(* IEC 61131-3 sources: plc-st-coding-agent/progress/evidence/f14_v14_remaining_20261113/jobs/custom_deepseek-v4pro, 30 files *)

(* ---- self-easy-01.candidate_01.st ---- *)
(*
ENGINEERING_CONTRACT
- activation: avgOut updates only when enable=TRUE AND avgEnable=TRUE AND count>0 after clipping count into 1..8.
- hold/retention: enable=FALSE, avgEnable=FALSE, or count<=0 leaves local_avg and avgOut unchanged this scan (S1/S2/S5).
- reset: none specified; avgOut persists until next valid compute; initial local_avg defaults to 0.0.
- boundary: count<=0 causes no division; count>8 uses first 8 samples only (PUB003/PUB004, no overflow).
- precision: sum accumulated in LINT, then converted to REAL and divided by REAL sample count (PUB005/PUB006).
- interface types preserved exactly; no edge-only triggers or interlocks added.
*)

(* CONTRACT_RULES [] *)

FUNCTION_BLOCK FB
VAR_INPUT
    enable: BOOL;
    values: ARRAY[1..8] OF INT;
    count: INT;
    avgEnable: BOOL;
END_VAR
VAR_OUTPUT
    avgOut: REAL;
END_VAR
VAR
    tmp_len: INT;
    tmp_sum: LINT;
    tmp_i: INT;
    local_avg: REAL := 0.0;
END_VAR

IF enable AND avgEnable THEN
    tmp_len := count;
    IF tmp_len < 0 THEN
        tmp_len := 0;
    END_IF;
    IF tmp_len > 8 THEN
        tmp_len := 8;
    END_IF;
    IF tmp_len > 0 THEN
        tmp_sum := 0;
        FOR tmp_i := 1 TO tmp_len BY 1 DO
            tmp_sum := tmp_sum + INT_TO_LINT(values[tmp_i]);
        END_FOR;
        local_avg := LINT_TO_REAL(tmp_sum) / INT_TO_REAL(tmp_len);
    END_IF;
END_IF;

avgOut := local_avg;

END_FUNCTION_BLOCK

(* ---- self-easy-01.raw_candidate_01.st ---- *)
(*
ENGINEERING_CONTRACT
- activation: avgOut updates only when enable=TRUE AND avgEnable=TRUE AND count>0 after clipping count into 1..8.
- hold/retention: enable=FALSE, avgEnable=FALSE, or count<=0 leaves local_avg and avgOut unchanged this scan (S1/S2/S5).
- reset: none specified; avgOut persists until next valid compute; initial local_avg defaults to 0.0.
- boundary: count<=0 causes no division; count>8 uses first 8 samples only (PUB003/PUB004, no overflow).
- precision: sum accumulated in LINT, then converted to REAL and divided by REAL sample count (PUB005/PUB006).
- interface types preserved exactly; no edge-only triggers or interlocks added.
*)

(* CONTRACT_RULES [] *)

FUNCTION_BLOCK FB
VAR_INPUT
    enable: BOOL;
    values: ARRAY[1..8] OF INT;
    count: INT;
    avgEnable: BOOL;
END_VAR
VAR_OUTPUT
    avgOut: REAL;
END_VAR
VAR
    tmp_len: INT;
    tmp_sum: LINT;
    tmp_i: INT;
    local_avg: REAL := 0.0;
END_VAR

IF enable AND avgEnable THEN
    tmp_len := count;
    IF tmp_len < 0 THEN
        tmp_len := 0;
    END_IF;
    IF tmp_len > 8 THEN
        tmp_len := 8;
    END_IF;
    IF tmp_len > 0 THEN
        tmp_sum := 0;
        FOR tmp_i := 1 TO tmp_len BY 1 DO
            tmp_sum := tmp_sum + INT_TO_LINT(values[tmp_i]);
        END_FOR;
        local_avg := LINT_TO_REAL(tmp_sum) / INT_TO_REAL(tmp_len);
    END_IF;
END_IF;

avgOut := local_avg;

END_FUNCTION_BLOCK

(* ---- self-easy-02.candidate_01.st ---- *)
FUNCTION_BLOCK FB
VAR_INPUT
    tankLevel : REAL;
    outletFlow : REAL;
    inletPermit : BOOL;
    resetBtn : BOOL;
END_VAR
VAR_OUTPUT
    pumpRun : BOOL;
    alarmHigh : BOOL;
    alarmLow : BOOL;
    outletValveOpen : BOOL;
END_VAR
VAR
    highLatched : BOOL := FALSE;
    lowLatched : BOOL := FALSE;
    prevResetBtn : BOOL := FALSE;
    tmp_resetRising : BOOL;
END_VAR

(* ENGINEERING_CONTRACT
   alarmHigh/alarmLow: set immediately at respective threshold, then latch.
   Activation: high >= 85.0, low <= 15.0 (REAL percent).
   Retention: remain latched when level returns to normal until reset.
   Reset: resetBtn rising edge clears each latch only if its danger is absent.
   Same-scan priority: danger condition overrides reset for the affected alarm.
   pumpRun: active only when inletPermit AND no alarm latched.
   outletValveOpen: inverse of low alarm; outletFlow is unused observation input.
*)

(* CONTRACT_RULES [] *)

tmp_resetRising := resetBtn AND NOT prevResetBtn;

IF tankLevel >= 85.0 THEN
    highLatched := TRUE;
ELSIF tmp_resetRising THEN
    highLatched := FALSE;
END_IF;

IF tankLevel <= 15.0 THEN
    lowLatched := TRUE;
ELSIF tmp_resetRising THEN
    lowLatched := FALSE;
END_IF;

alarmHigh := highLatched;
alarmLow := lowLatched;
pumpRun := inletPermit AND NOT highLatched AND NOT lowLatched;
outletValveOpen := NOT lowLatched;

prevResetBtn := resetBtn;

END_FUNCTION_BLOCK

(* ---- self-easy-02.raw_candidate_01.st ---- *)
FUNCTION_BLOCK FB
VAR_INPUT
    tankLevel : REAL;
    outletFlow : REAL;
    inletPermit : BOOL;
    resetBtn : BOOL;
END_VAR
VAR_OUTPUT
    pumpRun : BOOL;
    alarmHigh : BOOL;
    alarmLow : BOOL;
    outletValveOpen : BOOL;
END_VAR
VAR
    highLatched : BOOL := FALSE;
    lowLatched : BOOL := FALSE;
    prevResetBtn : BOOL := FALSE;
    tmp_resetRising : BOOL;
END_VAR

(* ENGINEERING_CONTRACT
   alarmHigh/alarmLow: set immediately at respective threshold, then latch.
   Activation: high >= 85.0, low <= 15.0 (REAL percent).
   Retention: remain latched when level returns to normal until reset.
   Reset: resetBtn rising edge clears each latch only if its danger is absent.
   Same-scan priority: danger condition overrides reset for the affected alarm.
   pumpRun: active only when inletPermit AND no alarm latched.
   outletValveOpen: inverse of low alarm; outletFlow is unused observation input.
*)

(* CONTRACT_RULES [] *)

tmp_resetRising := resetBtn AND NOT prevResetBtn;

IF tankLevel >= 85.0 THEN
    highLatched := TRUE;
ELSIF tmp_resetRising THEN
    highLatched := FALSE;
END_IF;

IF tankLevel <= 15.0 THEN
    lowLatched := TRUE;
ELSIF tmp_resetRising THEN
    lowLatched := FALSE;
END_IF;

alarmHigh := highLatched;
alarmLow := lowLatched;
pumpRun := inletPermit AND NOT highLatched AND NOT lowLatched;
outletValveOpen := NOT lowLatched;

prevResetBtn := resetBtn;

END_FUNCTION_BLOCK

(* ---- self-hard-01.candidate_01.st ---- *)
(*
ENGINEERING_CONTRACT
alarmActive: next = flowLow OR (prevActive AND !risingAck AND !(prevFlowLow AND prevAcked)).
  Retain on unacked condition loss; clear only when active-acked and flowLow drops, or ack rising while flowLow false.
alarmAcked: next = nextActive AND (!flowLow OR risingAck OR (prevFlowLow AND prevActive AND prevAcked)).
  True for active/acked or pending-clear; false when inactive or new flowLow after pending-clear.
highHigh = NOT sensorOK (combinational; no latch; auto clears same scan as sensorOK).
Memory: prevFlowLow/prevActive/prevAcked/prevAckBtn retained in VAR; update after output assignment.
Same-scan: risingAck computed before outputs; formulas use previous-cycle stored state; high priority independent.
Units: BOOL; no timers. See PUB001-PUB038.
*)
(* CONTRACT_RULES [] *)
FUNCTION_BLOCK FB
VAR_INPUT
    flowLow: BOOL;
    ackBtn: BOOL;
    sensorOK: BOOL;
END_VAR
VAR_OUTPUT
    alarmActive: BOOL;
    alarmAcked: BOOL;
    highHigh: BOOL;
END_VAR
VAR
    prevFlowLow: BOOL;
    prevAlarmActive: BOOL;
    prevAlarmAcked: BOOL;
    prevAckBtn: BOOL;
    risingAck: BOOL;
    nextActive: BOOL;
    nextAcked: BOOL;
    prevFlowLowAndAcked: BOOL;
    prevFlowLowActiveAcked: BOOL;
END_VAR

risingAck := ackBtn AND NOT prevAckBtn;

prevFlowLowAndAcked := prevFlowLow AND prevAlarmAcked;
prevFlowLowActiveAcked := prevFlowLow AND prevAlarmActive AND prevAlarmAcked;

nextActive := flowLow OR (prevAlarmActive AND NOT risingAck AND (NOT prevFlowLowAndAcked));
nextAcked := nextActive AND (NOT flowLow OR risingAck OR prevFlowLowActiveAcked);

alarmActive := nextActive;
alarmAcked := nextAcked;
highHigh := NOT sensorOK;

prevFlowLow := flowLow;
prevAlarmActive := nextActive;
prevAlarmAcked := nextAcked;
prevAckBtn := ackBtn;

END_FUNCTION_BLOCK

(* ---- self-hard-01.raw_candidate_01.st ---- *)
(*
ENGINEERING_CONTRACT
alarmActive: next = flowLow OR (prevActive AND !risingAck AND !(prevFlowLow AND prevAcked)).
  Retain on unacked condition loss; clear only when active-acked and flowLow drops, or ack rising while flowLow false.
alarmAcked: next = nextActive AND (!flowLow OR risingAck OR (prevFlowLow AND prevActive AND prevAcked)).
  True for active/acked or pending-clear; false when inactive or new flowLow after pending-clear.
highHigh = NOT sensorOK (combinational; no latch; auto clears same scan as sensorOK).
Memory: prevFlowLow/prevActive/prevAcked/prevAckBtn retained in VAR; update after output assignment.
Same-scan: risingAck computed before outputs; formulas use previous-cycle stored state; high priority independent.
Units: BOOL; no timers. See PUB001-PUB038.
*)
(* CONTRACT_RULES [] *)
FUNCTION_BLOCK FB
VAR_INPUT
    flowLow: BOOL;
    ackBtn: BOOL;
    sensorOK: BOOL;
END_VAR
VAR_OUTPUT
    alarmActive: BOOL;
    alarmAcked: BOOL;
    highHigh: BOOL;
END_VAR
VAR
    prevFlowLow: BOOL;
    prevAlarmActive: BOOL;
    prevAlarmAcked: BOOL;
    prevAckBtn: BOOL;
    risingAck: BOOL;
    nextActive: BOOL;
    nextAcked: BOOL;
    prevFlowLowAndAcked: BOOL;
    prevFlowLowActiveAcked: BOOL;
END_VAR

risingAck := ackBtn AND NOT prevAckBtn;

prevFlowLowAndAcked := prevFlowLow AND prevAlarmAcked;
prevFlowLowActiveAcked := prevFlowLow AND prevAlarmActive AND prevAlarmAcked;

nextActive := flowLow OR (prevAlarmActive AND NOT risingAck AND (NOT prevFlowLowAndAcked));
nextAcked := nextActive AND (NOT flowLow OR risingAck OR prevFlowLowActiveAcked);

alarmActive := nextActive;
alarmAcked := nextAcked;
highHigh := NOT sensorOK;

prevFlowLow := flowLow;
prevAlarmActive := nextActive;
prevAlarmAcked := nextAcked;
prevAckBtn := ackBtn;

END_FUNCTION_BLOCK

(* ---- self-hard-02.candidate_01.st ---- *)
FUNCTION_BLOCK FB
VAR_INPUT
    startBtn : BOOL;
    abortBtn : BOOL;
    setpoint : REAL;
    pv : REAL;
    maxDuration : INT;
END_VAR
VAR_OUTPUT
    elapsed : INT;
    phase : INT;
    timeout : BOOL;
END_VAR
VAR
    prevStartBtn : BOOL;
    tmpStartRising : BOOL;
    tmpPrevPhase : INT;
    tmpPrevElapsed : INT;
    tmpPrevTimeout : BOOL;
    tmpIsRunPrev : BOOL;
    tmpNewElapsed : INT;
END_VAR

(* ENGINEERING_CONTRACT
   phase: 0 idle, 1 heating, 2 soaking, 3 done, 9 aborted.
   Activation: phase=1 on start rising without abort; phase=2 when previous run phase is 1 and pv>=setpoint before timeout; phase=3 when elapsed>=maxDuration; phase=9 on abort.
   Retention: phase 3/9 hold until new start or abort; start resets to 1 and clears elapsed/timeout; abort from 3/9 preserves elapsed/timeout.
   elapsed: counts scans when previous phase is 1 or 2 and no abort/start rising. Reset to 0 on start; frozen in 3/9; frozen on abort.
   timeout: set TRUE when new elapsed>=maxDuration (scan count); cleared on start; frozen on abort; otherwise equals timeout condition.
   Priority: abort > start rising > running count; same-scan start edge consumed even under abort.
   Units: elapsed/maxDuration in scan counts, INT; no timer used.
*)

(* CONTRACT_RULES [] *)

tmpStartRising := startBtn AND NOT prevStartBtn;
tmpPrevPhase := phase;
tmpPrevElapsed := elapsed;
tmpPrevTimeout := timeout;
tmpIsRunPrev := (tmpPrevPhase = 1) OR (tmpPrevPhase = 2);

IF abortBtn THEN
    phase := 9;
    elapsed := tmpPrevElapsed;
    timeout := tmpPrevTimeout;
ELSIF tmpStartRising THEN
    phase := 1;
    elapsed := 0;
    timeout := FALSE;
ELSE
    IF tmpIsRunPrev THEN
        tmpNewElapsed := tmpPrevElapsed + 1;
        elapsed := tmpNewElapsed;
        IF tmpNewElapsed >= maxDuration THEN
            timeout := TRUE;
            phase := 3;
        ELSE
            timeout := FALSE;
            IF tmpPrevPhase = 2 THEN
                phase := 2;
            ELSE
                IF pv >= setpoint THEN
                    phase := 2;
                ELSE
                    phase := 1;
                END_IF;
            END_IF;
        END_IF;
    ELSE
        phase := tmpPrevPhase;
        elapsed := tmpPrevElapsed;
        timeout := tmpPrevTimeout;
    END_IF;
END_IF;

prevStartBtn := startBtn;
END_FUNCTION_BLOCK

(* ---- self-hard-02.raw_candidate_01.st ---- *)
FUNCTION_BLOCK FB
VAR_INPUT
    startBtn : BOOL;
    abortBtn : BOOL;
    setpoint : REAL;
    pv : REAL;
    maxDuration : INT;
END_VAR
VAR_OUTPUT
    elapsed : INT;
    phase : INT;
    timeout : BOOL;
END_VAR
VAR
    prevStartBtn : BOOL;
    tmpStartRising : BOOL;
    tmpPrevPhase : INT;
    tmpPrevElapsed : INT;
    tmpPrevTimeout : BOOL;
    tmpIsRunPrev : BOOL;
    tmpNewElapsed : INT;
END_VAR

(* ENGINEERING_CONTRACT
   phase: 0 idle, 1 heating, 2 soaking, 3 done, 9 aborted.
   Activation: phase=1 on start rising without abort; phase=2 when previous run phase is 1 and pv>=setpoint before timeout; phase=3 when elapsed>=maxDuration; phase=9 on abort.
   Retention: phase 3/9 hold until new start or abort; start resets to 1 and clears elapsed/timeout; abort from 3/9 preserves elapsed/timeout.
   elapsed: counts scans when previous phase is 1 or 2 and no abort/start rising. Reset to 0 on start; frozen in 3/9; frozen on abort.
   timeout: set TRUE when new elapsed>=maxDuration (scan count); cleared on start; frozen on abort; otherwise equals timeout condition.
   Priority: abort > start rising > running count; same-scan start edge consumed even under abort.
   Units: elapsed/maxDuration in scan counts, INT; no timer used.
*)

(* CONTRACT_RULES [] *)

tmpStartRising := startBtn AND NOT prevStartBtn;
tmpPrevPhase := phase;
tmpPrevElapsed := elapsed;
tmpPrevTimeout := timeout;
tmpIsRunPrev := (tmpPrevPhase = 1) OR (tmpPrevPhase = 2);

IF abortBtn THEN
    phase := 9;
    elapsed := tmpPrevElapsed;
    timeout := tmpPrevTimeout;
ELSIF tmpStartRising THEN
    phase := 1;
    elapsed := 0;
    timeout := FALSE;
ELSE
    IF tmpIsRunPrev THEN
        tmpNewElapsed := tmpPrevElapsed + 1;
        elapsed := tmpNewElapsed;
        IF tmpNewElapsed >= maxDuration THEN
            timeout := TRUE;
            phase := 3;
        ELSE
            timeout := FALSE;
            IF tmpPrevPhase = 2 THEN
                phase := 2;
            ELSE
                IF pv >= setpoint THEN
                    phase := 2;
                ELSE
                    phase := 1;
                END_IF;
            END_IF;
        END_IF;
    ELSE
        phase := tmpPrevPhase;
        elapsed := tmpPrevElapsed;
        timeout := tmpPrevTimeout;
    END_IF;
END_IF;

prevStartBtn := startBtn;
END_FUNCTION_BLOCK

(* ---- self-hard-03.candidate_01.st ---- *)
(* ENGINEERING_CONTRACT
   count: updated by successful pop then successful push; retained otherwise; initial 0; bounds 0..8; S1,S6.
   full: combinational = (count=8); no latch; S1.
   empty: combinational = (count=0); no latch; S1.
   head: count=0 -> 0; else fifo[1]; combinational after actions; S5.
   fifo valid prefix: compact; shift on successful pop; append on successful push; S4,S7,S8.
   Edge history: local_push_prev/local_pop_prev retained; initial FALSE; updated each scan.
   Priority: pop rising executes before push rising; capacity checked after pop; PUB requirement order.
*)
(* CONTRACT_RULES [] *)
FUNCTION_BLOCK FB
VAR_INPUT
    pushEn : BOOL;
    pushItem : INT;
    popEn : BOOL;
END_VAR
VAR_OUTPUT
    count : INT;
    full : BOOL;
    empty : BOOL;
    head : INT;
END_VAR
VAR_IN_OUT
    fifo : ARRAY[1..8] OF INT;
END_VAR
VAR
    local_push_prev : BOOL := FALSE;
    local_pop_prev : BOOL := FALSE;
    local_count : INT := 0;
    local_rising_push : BOOL;
    local_rising_pop : BOOL;
    i : INT;
END_VAR

(* 计算上升沿，历史在扫描结束时更新 *)
local_rising_push := pushEn AND NOT local_push_prev;
local_rising_pop := popEn AND NOT local_pop_prev;

(* 先执行出队 *)
IF local_rising_pop AND (local_count > 0) THEN
    IF local_count > 1 THEN
        FOR i := 1 TO local_count - 1 DO
            fifo[i] := fifo[i + 1];
        END_FOR;
    END_IF;
    local_count := local_count - 1;
END_IF;

(* 后执行入队 *)
IF local_rising_push AND (local_count < 8) THEN
    local_count := local_count + 1;
    fifo[local_count] := pushItem;
END_IF;

(* 输出 *)
count := local_count;
full := (local_count = 8);
empty := (local_count = 0);
IF local_count = 0 THEN
    head := 0;
ELSE
    head := fifo[1];
END_IF;

(* 更新输入历史 *)
local_push_prev := pushEn;
local_pop_prev := popEn;

END_FUNCTION_BLOCK

(* ---- self-hard-03.raw_candidate_01.st ---- *)
(* ENGINEERING_CONTRACT
   count: updated by successful pop then successful push; retained otherwise; initial 0; bounds 0..8; S1,S6.
   full: combinational = (count=8); no latch; S1.
   empty: combinational = (count=0); no latch; S1.
   head: count=0 -> 0; else fifo[1]; combinational after actions; S5.
   fifo valid prefix: compact; shift on successful pop; append on successful push; S4,S7,S8.
   Edge history: local_push_prev/local_pop_prev retained; initial FALSE; updated each scan.
   Priority: pop rising executes before push rising; capacity checked after pop; PUB requirement order.
*)
(* CONTRACT_RULES [] *)
FUNCTION_BLOCK FB
VAR_INPUT
    pushEn : BOOL;
    pushItem : INT;
    popEn : BOOL;
END_VAR
VAR_OUTPUT
    count : INT;
    full : BOOL;
    empty : BOOL;
    head : INT;
END_VAR
VAR_IN_OUT
    fifo : ARRAY[1..8] OF INT;
END_VAR
VAR
    local_push_prev : BOOL := FALSE;
    local_pop_prev : BOOL := FALSE;
    local_count : INT := 0;
    local_rising_push : BOOL;
    local_rising_pop : BOOL;
    i : INT;
END_VAR

(* 计算上升沿，历史在扫描结束时更新 *)
local_rising_push := pushEn AND NOT local_push_prev;
local_rising_pop := popEn AND NOT local_pop_prev;

(* 先执行出队 *)
IF local_rising_pop AND (local_count > 0) THEN
    IF local_count > 1 THEN
        FOR i := 1 TO local_count - 1 DO
            fifo[i] := fifo[i + 1];
        END_FOR;
    END_IF;
    local_count := local_count - 1;
END_IF;

(* 后执行入队 *)
IF local_rising_push AND (local_count < 8) THEN
    local_count := local_count + 1;
    fifo[local_count] := pushItem;
END_IF;

(* 输出 *)
count := local_count;
full := (local_count = 8);
empty := (local_count = 0);
IF local_count = 0 THEN
    head := 0;
ELSE
    head := fifo[1];
END_IF;

(* 更新输入历史 *)
local_push_prev := pushEn;
local_pop_prev := popEn;

END_FUNCTION_BLOCK

(* ---- self-hard-04.candidate_01.st ---- *)
(* ENGINEERING_CONTRACT
  runningCount: combinational; activation every scan; clip demand to 0..5; no retention/reset; same-scan priority: computed first; range 0..5 [PUB001,S1].
  leadPump: stored selection; activation: positive demand with prevLead=0 -> global (hours,pump) min (tie smallest pump); positive prevLead valid + rotated TRUE and oldLeadHours-globalMinHours > 50 -> global min; else retain; deactivation/reset: demand<=0 -> 0; units 1..5,0=none [PUB004,S2,S3,S6,S7].
  lagPump: stored selection; activation/update: demand>=2 and (lead changed OR clipped demand rose) -> min among pumps excluding current lead (tie smallest pump); retention: otherwise while demand>=2; deactivation/reset: demand<=1 -> 0; units 1..5,0=none [PUB005,S8,S9].
  Arrays accessed with indices 1..5 only; previous outputs kept in static VAR [PUB006].
*)
(* CONTRACT_RULES [] *)
FUNCTION_BLOCK FB
VAR_INPUT
    demand : INT;
    runHours : ARRAY[1..5] OF LINT;
    rotated : BOOL;
END_VAR
VAR_OUTPUT
    leadPump : INT;
    lagPump : INT;
    runningCount : INT;
END_VAR
VAR
    local_prevLeadPump : INT := 0;
    local_prevLagPump : INT := 0;
    local_prevRunningCount : INT := 0;
    local_demandClipped : INT;
    local_i : INT;
    local_minPumpAll : INT;
    local_minHoursAll : LINT;
    local_minPumpExcl : INT;
    local_minHoursExcl : LINT;
    local_firstFound : BOOL;
END_VAR

IF demand < 0 THEN
    local_demandClipped := 0;
ELSIF demand > 5 THEN
    local_demandClipped := 5;
ELSE
    local_demandClipped := demand;
END_IF;

runningCount := local_demandClipped;

IF local_demandClipped <= 0 THEN
    leadPump := 0;
    lagPump := 0;
ELSE
    local_minPumpAll := 1;
    local_minHoursAll := runHours[1];
    FOR local_i := 2 TO 5 DO
        IF (runHours[local_i] < local_minHoursAll) OR
           ((runHours[local_i] = local_minHoursAll) AND (local_i < local_minPumpAll)) THEN
            local_minPumpAll := local_i;
            local_minHoursAll := runHours[local_i];
        END_IF;
    END_FOR;

    IF local_prevLeadPump = 0 THEN
        leadPump := local_minPumpAll;
    ELSE
        leadPump := local_prevLeadPump;
        IF rotated THEN
            IF runHours[local_prevLeadPump] - local_minHoursAll > LINT#50 THEN
                leadPump := local_minPumpAll;
            END_IF;
        END_IF;
    END_IF;

    IF local_demandClipped = 1 THEN
        lagPump := 0;
    ELSE
        IF (leadPump <> local_prevLeadPump) OR (local_demandClipped > local_prevRunningCount) THEN
            local_minPumpExcl := 0;
            local_minHoursExcl := 0;
            local_firstFound := FALSE;
            FOR local_i := 1 TO 5 DO
                IF local_i <> leadPump THEN
                    IF NOT local_firstFound THEN
                        local_minPumpExcl := local_i;
                        local_minHoursExcl := runHours[local_i];
                        local_firstFound := TRUE;
                    ELSE
                        IF (runHours[local_i] < local_minHoursExcl) OR
                           ((runHours[local_i] = local_minHoursExcl) AND (local_i < local_minPumpExcl)) THEN
                            local_minPumpExcl := local_i;
                            local_minHoursExcl := runHours[local_i];
                        END_IF;
                    END_IF;
                END_IF;
            END_FOR;
            lagPump := local_minPumpExcl;
        ELSE
            lagPump := local_prevLagPump;
        END_IF;
    END_IF;
END_IF;

local_prevLeadPump := leadPump;
local_prevLagPump := lagPump;
local_prevRunningCount := runningCount;

END_FUNCTION_BLOCK

(* ---- self-hard-04.raw_candidate_01.st ---- *)
(* ENGINEERING_CONTRACT
  runningCount: combinational; activation every scan; clip demand to 0..5; no retention/reset; same-scan priority: computed first; range 0..5 [PUB001,S1].
  leadPump: stored selection; activation: positive demand with prevLead=0 -> global (hours,pump) min (tie smallest pump); positive prevLead valid + rotated TRUE and oldLeadHours-globalMinHours > 50 -> global min; else retain; deactivation/reset: demand<=0 -> 0; units 1..5,0=none [PUB004,S2,S3,S6,S7].
  lagPump: stored selection; activation/update: demand>=2 and (lead changed OR clipped demand rose) -> min among pumps excluding current lead (tie smallest pump); retention: otherwise while demand>=2; deactivation/reset: demand<=1 -> 0; units 1..5,0=none [PUB005,S8,S9].
  Arrays accessed with indices 1..5 only; previous outputs kept in static VAR [PUB006].
*)
(* CONTRACT_RULES [] *)
FUNCTION_BLOCK FB
VAR_INPUT
    demand : INT;
    runHours : ARRAY[1..5] OF LINT;
    rotated : BOOL;
END_VAR
VAR_OUTPUT
    leadPump : INT;
    lagPump : INT;
    runningCount : INT;
END_VAR
VAR
    local_prevLeadPump : INT := 0;
    local_prevLagPump : INT := 0;
    local_prevRunningCount : INT := 0;
    local_demandClipped : INT;
    local_i : INT;
    local_minPumpAll : INT;
    local_minHoursAll : LINT;
    local_minPumpExcl : INT;
    local_minHoursExcl : LINT;
    local_firstFound : BOOL;
END_VAR

IF demand < 0 THEN
    local_demandClipped := 0;
ELSIF demand > 5 THEN
    local_demandClipped := 5;
ELSE
    local_demandClipped := demand;
END_IF;

runningCount := local_demandClipped;

IF local_demandClipped <= 0 THEN
    leadPump := 0;
    lagPump := 0;
ELSE
    local_minPumpAll := 1;
    local_minHoursAll := runHours[1];
    FOR local_i := 2 TO 5 DO
        IF (runHours[local_i] < local_minHoursAll) OR
           ((runHours[local_i] = local_minHoursAll) AND (local_i < local_minPumpAll)) THEN
            local_minPumpAll := local_i;
            local_minHoursAll := runHours[local_i];
        END_IF;
    END_FOR;

    IF local_prevLeadPump = 0 THEN
        leadPump := local_minPumpAll;
    ELSE
        leadPump := local_prevLeadPump;
        IF rotated THEN
            IF runHours[local_prevLeadPump] - local_minHoursAll > LINT#50 THEN
                leadPump := local_minPumpAll;
            END_IF;
        END_IF;
    END_IF;

    IF local_demandClipped = 1 THEN
        lagPump := 0;
    ELSE
        IF (leadPump <> local_prevLeadPump) OR (local_demandClipped > local_prevRunningCount) THEN
            local_minPumpExcl := 0;
            local_minHoursExcl := 0;
            local_firstFound := FALSE;
            FOR local_i := 1 TO 5 DO
                IF local_i <> leadPump THEN
                    IF NOT local_firstFound THEN
                        local_minPumpExcl := local_i;
                        local_minHoursExcl := runHours[local_i];
                        local_firstFound := TRUE;
                    ELSE
                        IF (runHours[local_i] < local_minHoursExcl) OR
                           ((runHours[local_i] = local_minHoursExcl) AND (local_i < local_minPumpExcl)) THEN
                            local_minPumpExcl := local_i;
                            local_minHoursExcl := runHours[local_i];
                        END_IF;
                    END_IF;
                END_IF;
            END_FOR;
            lagPump := local_minPumpExcl;
        ELSE
            lagPump := local_prevLagPump;
        END_IF;
    END_IF;
END_IF;

local_prevLeadPump := leadPump;
local_prevLagPump := lagPump;
local_prevRunningCount := runningCount;

END_FUNCTION_BLOCK

(* ---- self-hard-05.candidate_01.st ---- *)
(* ENGINEERING_CONTRACT
tripLatched: set same scan when runRequest=TRUE AND flameOK=FALSE; held; clear only on rising resetBtn while runRequest=FALSE AND flameOK=FALSE; fire-set dominates. PUB001 PUB006 PUB030 PUB031 PUB059.
fuelPermit: combinational = runRequest AND flameOK AND NOT tripLatched. PUB005 PUB060.
o2Fault: combinational = NOT o2Valid OR o2PV<0.0 OR o2PV>21.0. PUB012 PUB061.
trimEnable: combinational = fuelPermit AND NOT o2Fault. PUB008 PUB061.
airTrim: if trimEnable then clamp(2.0*(2.0-o2PV), -10.0, 10.0) else 0.0; saturation reaches -10 only when o2PV>7.0. PUB010 PUB011 PUB014 PUB015 PUB052 PUB053.
airCommand: if fuelPermit then clamp(baseAir+airTrim, 0.0, 100.0) else 0.0. PUB011 PUB013 PUB015 PUB045 PUB046 PUB055.
reset edge: detected once per scan via prevResetBtn; no timer. Units: REAL %, BOOL, scan cycle. PUB006 PUB030 PUB031.
*)
(* CONTRACT_RULES [] *)
FUNCTION_BLOCK FB
VAR_INPUT
    runRequest : BOOL;
    flameOK : BOOL;
    o2Valid : BOOL;
    o2PV : REAL;
    baseAir : REAL;
    resetBtn : BOOL;
END_VAR
VAR_OUTPUT
    fuelPermit : BOOL;
    trimEnable : BOOL;
    airTrim : REAL;
    airCommand : REAL;
    tripLatched : BOOL;
    o2Fault : BOOL;
END_VAR
VAR
    prevResetBtn : BOOL := FALSE;
    tmp_resetRise : BOOL;
    tmp_prevTrip : BOOL;
    tmp_rawTrim : REAL;
    tmp_sum : REAL;
END_VAR

    tmp_resetRise := resetBtn AND NOT prevResetBtn;
    tmp_prevTrip := tripLatched;
    tripLatched := (runRequest AND NOT flameOK)
                   OR (tmp_prevTrip AND NOT (tmp_resetRise AND NOT runRequest AND NOT flameOK));
    prevResetBtn := resetBtn;

    fuelPermit := runRequest AND flameOK AND NOT tripLatched;

    o2Fault := (NOT o2Valid) OR (o2PV < 0.0) OR (o2PV > 21.0);
    trimEnable := fuelPermit AND NOT o2Fault;

    IF trimEnable THEN
        tmp_rawTrim := 2.0 * (2.0 - o2PV);
        IF tmp_rawTrim < -10.0 THEN
            airTrim := -10.0;
        ELSIF tmp_rawTrim > 10.0 THEN
            airTrim := 10.0;
        ELSE
            airTrim := tmp_rawTrim;
        END_IF;
    ELSE
        airTrim := 0.0;
    END_IF;

    IF fuelPermit THEN
        tmp_sum := baseAir + airTrim;
        IF tmp_sum < 0.0 THEN
            airCommand := 0.0;
        ELSIF tmp_sum > 100.0 THEN
            airCommand := 100.0;
        ELSE
            airCommand := tmp_sum;
        END_IF;
    ELSE
        airCommand := 0.0;
    END_IF;

END_FUNCTION_BLOCK

(* ---- self-hard-05.raw_candidate_01.st ---- *)
(* ENGINEERING_CONTRACT
tripLatched: set same scan when runRequest=TRUE AND flameOK=FALSE; held; clear only on rising resetBtn while runRequest=FALSE AND flameOK=FALSE; fire-set dominates. PUB001 PUB006 PUB030 PUB031 PUB059.
fuelPermit: combinational = runRequest AND flameOK AND NOT tripLatched. PUB005 PUB060.
o2Fault: combinational = NOT o2Valid OR o2PV<0.0 OR o2PV>21.0. PUB012 PUB061.
trimEnable: combinational = fuelPermit AND NOT o2Fault. PUB008 PUB061.
airTrim: if trimEnable then clamp(2.0*(2.0-o2PV), -10.0, 10.0) else 0.0; saturation reaches -10 only when o2PV>7.0. PUB010 PUB011 PUB014 PUB015 PUB052 PUB053.
airCommand: if fuelPermit then clamp(baseAir+airTrim, 0.0, 100.0) else 0.0. PUB011 PUB013 PUB015 PUB045 PUB046 PUB055.
reset edge: detected once per scan via prevResetBtn; no timer. Units: REAL %, BOOL, scan cycle. PUB006 PUB030 PUB031.
*)
(* CONTRACT_RULES [] *)
FUNCTION_BLOCK FB
VAR_INPUT
    runRequest : BOOL;
    flameOK : BOOL;
    o2Valid : BOOL;
    o2PV : REAL;
    baseAir : REAL;
    resetBtn : BOOL;
END_VAR
VAR_OUTPUT
    fuelPermit : BOOL;
    trimEnable : BOOL;
    airTrim : REAL;
    airCommand : REAL;
    tripLatched : BOOL;
    o2Fault : BOOL;
END_VAR
VAR
    prevResetBtn : BOOL := FALSE;
    tmp_resetRise : BOOL;
    tmp_prevTrip : BOOL;
    tmp_rawTrim : REAL;
    tmp_sum : REAL;
END_VAR

    tmp_resetRise := resetBtn AND NOT prevResetBtn;
    tmp_prevTrip := tripLatched;
    tripLatched := (runRequest AND NOT flameOK)
                   OR (tmp_prevTrip AND NOT (tmp_resetRise AND NOT runRequest AND NOT flameOK));
    prevResetBtn := resetBtn;

    fuelPermit := runRequest AND flameOK AND NOT tripLatched;

    o2Fault := (NOT o2Valid) OR (o2PV < 0.0) OR (o2PV > 21.0);
    trimEnable := fuelPermit AND NOT o2Fault;

    IF trimEnable THEN
        tmp_rawTrim := 2.0 * (2.0 - o2PV);
        IF tmp_rawTrim < -10.0 THEN
            airTrim := -10.0;
        ELSIF tmp_rawTrim > 10.0 THEN
            airTrim := 10.0;
        ELSE
            airTrim := tmp_rawTrim;
        END_IF;
    ELSE
        airTrim := 0.0;
    END_IF;

    IF fuelPermit THEN
        tmp_sum := baseAir + airTrim;
        IF tmp_sum < 0.0 THEN
            airCommand := 0.0;
        ELSIF tmp_sum > 100.0 THEN
            airCommand := 100.0;
        ELSE
            airCommand := tmp_sum;
        END_IF;
    ELSE
        airCommand := 0.0;
    END_IF;

END_FUNCTION_BLOCK

(* ---- self-hard-06.candidate_01.st ---- *)
(* ENGINEERING_CONTRACT
  tripLatched: active same scan on trip condition (run & !pressureValid) OR (run & pressureValid & pressure>=4500.0);
               retains until legal reset edge: resetBtn rising & !run & pressureValid & pressure<=4200.0.
  fuelPermit: combinational = run & !tripLatched, evaluated after latch update.
  currentCauseMask: low nibble recalculated each scan; !run=0, invalid=1, valid overpressure evaluates stuck/excess/unlocated, below 4500=0.
  latchedCauseMask: OR currentCauseMask while tripLatched; clear when !tripLatched; low 4 bits only.
  stuckCounter: counts consecutive full overpressure+valve-condition scans; reset on any interruption.
  diagnosticActive: currentCauseMask<>0.
  Unspecified: scan period undefined; initial resetBtn edge state considered FALSE.
*)
(* CONTRACT_RULES [] *)
FUNCTION_BLOCK FB
VAR_INPUT
    runRequest : BOOL;
    pressure : REAL;
    pressureValid : BOOL;
    fuelFlow : REAL;
    steamFlow : REAL;
    outletCmd : INT;
    outletFeedback : INT;
    resetBtn : BOOL;
END_VAR
VAR_OUTPUT
    tripLatched : BOOL;
    fuelPermit : BOOL;
    currentCauseMask : WORD;
    latchedCauseMask : WORD;
    diagnosticActive : BOOL;
END_VAR
VAR
    lastResetBtn : BOOL := FALSE;
    stuckCounter : INT := 0;
    tmp_resetRising : BOOL;
    tmp_overpressure : BOOL;
    tmp_invalid : BOOL;
    tmp_tripCondition : BOOL;
    tmp_legalReset : BOOL;
    tmp_stuckCond : BOOL;
    tmp_stuckBit : BOOL;
    tmp_excessBit : BOOL;
END_VAR

tmp_resetRising := resetBtn AND NOT lastResetBtn;
lastResetBtn := resetBtn;

tmp_overpressure := runRequest AND pressureValid AND pressure >= 4500.0;
tmp_invalid := runRequest AND NOT pressureValid;
tmp_tripCondition := tmp_overpressure OR tmp_invalid;
tmp_legalReset := tmp_resetRising AND NOT runRequest AND pressureValid AND pressure <= 4200.0;

IF NOT runRequest THEN
    currentCauseMask := WORD#0;
    stuckCounter := 0;
ELSIF NOT pressureValid THEN
    currentCauseMask := WORD#1;
    stuckCounter := 0;
ELSIF pressure >= 4500.0 THEN
    tmp_stuckCond := (outletCmd >= 50) AND (outletFeedback <= 10);
    IF tmp_stuckCond THEN
        stuckCounter := stuckCounter + 1;
    ELSE
        stuckCounter := 0;
    END_IF;
    tmp_stuckBit := stuckCounter >= 3;
    tmp_excessBit := (fuelFlow >= 4.0) AND (steamFlow <= 10.0);
    IF tmp_stuckBit AND tmp_excessBit THEN
        currentCauseMask := WORD#6;
    ELSIF tmp_excessBit THEN
        currentCauseMask := WORD#4;
    ELSIF tmp_stuckBit THEN
        currentCauseMask := WORD#2;
    ELSE
        currentCauseMask := WORD#8;
    END_IF;
ELSE
    currentCauseMask := WORD#0;
    stuckCounter := 0;
END_IF;

IF tmp_tripCondition THEN
    tripLatched := TRUE;
ELSIF tmp_legalReset THEN
    tripLatched := FALSE;
END_IF;

IF tripLatched THEN
    latchedCauseMask := (latchedCauseMask OR currentCauseMask) AND WORD#15;
ELSE
    latchedCauseMask := WORD#0;
END_IF;

fuelPermit := runRequest AND NOT tripLatched;
diagnosticActive := currentCauseMask <> WORD#0;

END_FUNCTION_BLOCK

(* ---- self-hard-06.raw_candidate_01.st ---- *)
(* ENGINEERING_CONTRACT
  tripLatched: active same scan on trip condition (run & !pressureValid) OR (run & pressureValid & pressure>=4500.0);
               retains until legal reset edge: resetBtn rising & !run & pressureValid & pressure<=4200.0.
  fuelPermit: combinational = run & !tripLatched, evaluated after latch update.
  currentCauseMask: low nibble recalculated each scan; !run=0, invalid=1, valid overpressure evaluates stuck/excess/unlocated, below 4500=0.
  latchedCauseMask: OR currentCauseMask while tripLatched; clear when !tripLatched; low 4 bits only.
  stuckCounter: counts consecutive full overpressure+valve-condition scans; reset on any interruption.
  diagnosticActive: currentCauseMask<>0.
  Unspecified: scan period undefined; initial resetBtn edge state considered FALSE.
*)
(* CONTRACT_RULES [] *)
FUNCTION_BLOCK FB
VAR_INPUT
    runRequest : BOOL;
    pressure : REAL;
    pressureValid : BOOL;
    fuelFlow : REAL;
    steamFlow : REAL;
    outletCmd : INT;
    outletFeedback : INT;
    resetBtn : BOOL;
END_VAR
VAR_OUTPUT
    tripLatched : BOOL;
    fuelPermit : BOOL;
    currentCauseMask : WORD;
    latchedCauseMask : WORD;
    diagnosticActive : BOOL;
END_VAR
VAR
    lastResetBtn : BOOL := FALSE;
    stuckCounter : INT := 0;
    tmp_resetRising : BOOL;
    tmp_overpressure : BOOL;
    tmp_invalid : BOOL;
    tmp_tripCondition : BOOL;
    tmp_legalReset : BOOL;
    tmp_stuckCond : BOOL;
    tmp_stuckBit : BOOL;
    tmp_excessBit : BOOL;
END_VAR

tmp_resetRising := resetBtn AND NOT lastResetBtn;
lastResetBtn := resetBtn;

tmp_overpressure := runRequest AND pressureValid AND pressure >= 4500.0;
tmp_invalid := runRequest AND NOT pressureValid;
tmp_tripCondition := tmp_overpressure OR tmp_invalid;
tmp_legalReset := tmp_resetRising AND NOT runRequest AND pressureValid AND pressure <= 4200.0;

IF NOT runRequest THEN
    currentCauseMask := WORD#0;
    stuckCounter := 0;
ELSIF NOT pressureValid THEN
    currentCauseMask := WORD#1;
    stuckCounter := 0;
ELSIF pressure >= 4500.0 THEN
    tmp_stuckCond := (outletCmd >= 50) AND (outletFeedback <= 10);
    IF tmp_stuckCond THEN
        stuckCounter := stuckCounter + 1;
    ELSE
        stuckCounter := 0;
    END_IF;
    tmp_stuckBit := stuckCounter >= 3;
    tmp_excessBit := (fuelFlow >= 4.0) AND (steamFlow <= 10.0);
    IF tmp_stuckBit AND tmp_excessBit THEN
        currentCauseMask := WORD#6;
    ELSIF tmp_excessBit THEN
        currentCauseMask := WORD#4;
    ELSIF tmp_stuckBit THEN
        currentCauseMask := WORD#2;
    ELSE
        currentCauseMask := WORD#8;
    END_IF;
ELSE
    currentCauseMask := WORD#0;
    stuckCounter := 0;
END_IF;

IF tmp_tripCondition THEN
    tripLatched := TRUE;
ELSIF tmp_legalReset THEN
    tripLatched := FALSE;
END_IF;

IF tripLatched THEN
    latchedCauseMask := (latchedCauseMask OR currentCauseMask) AND WORD#15;
ELSE
    latchedCauseMask := WORD#0;
END_IF;

fuelPermit := runRequest AND NOT tripLatched;
diagnosticActive := currentCauseMask <> WORD#0;

END_FUNCTION_BLOCK

(* ---- self-hard-07.candidate_01.st ---- *)
FUNCTION_BLOCK FB
VAR_INPUT
    mode : INT;
    resetBtn : BOOL;
    scanSeconds : REAL;
    tempSP : REAL;
    tempPV : REAL;
    flowPV : REAL;
    manualFlowSP : REAL;
    manualValve : REAL;
END_VAR
VAR_OUTPUT
    flowSP : REAL;
    valveCommand : REAL;
    fault : BOOL;
    normalMode : BOOL;
END_VAR
VAR
    first : BOOL := TRUE;
    prevMode : INT := 0;
    prevResetBtn : BOOL := FALSE;
    prevFlowSP : REAL := 0.0;
    prevValveCmd : REAL := 0.0;
    accT : REAL := 0.0;
    accF : REAL := 0.0;
    tmp_eT : REAL;
    tmp_eF : REAL;
    tmp_flowUnlim : REAL;
    tmp_valveUnlim : REAL;
    tmp_resetRising : BOOL;
    tmp_modeChanged : BOOL;
END_VAR

(* ENGINEERING_CONTRACT
   flowSP: manual/limited PI output; retained via prevFlowSP between scans; reset/fault/switch presets.
   valveCommand: manual/limited PI output; retained via prevValveCmd; reset/fault/switch presets.
   fault: combinational from mode/scanSeconds; no latch.
   normalMode: true only in stable valid mode with no first/reset/fault/mode change.
   Reset rising: outputs=manual values, integrators preloaded; fault still reports current mode/scanSeconds.
   PI back-calculates accT/accF from final outputs every scan, preventing integral windup.
   Units: flowSP t/h, valveCommand %, accT t/h, accF %, scanSeconds s. PUB001-PUB065.
*)
(* CONTRACT_RULES [] *)

fault := (mode < 0) OR (mode > 2) OR (scanSeconds <= 0.0) OR (scanSeconds > 10.0);
tmp_resetRising := resetBtn AND NOT prevResetBtn;
normalMode := FALSE;

IF first THEN
    flowSP := manualFlowSP;
    valveCommand := manualValve;
ELSIF fault THEN
    flowSP := manualFlowSP;
    valveCommand := manualValve;
ELSIF tmp_resetRising THEN
    flowSP := manualFlowSP;
    valveCommand := manualValve;
ELSE
    tmp_modeChanged := (mode <> prevMode);
    IF tmp_modeChanged THEN
        IF mode = 2 THEN
            flowSP := prevFlowSP;
            valveCommand := prevValveCmd;
        ELSE
            flowSP := manualFlowSP;
            valveCommand := prevValveCmd;
        END_IF;
    ELSE
        normalMode := TRUE;
        CASE mode OF
            0:
                flowSP := manualFlowSP;
                valveCommand := manualValve;

            1:
                flowSP := manualFlowSP;
                tmp_eF := flowSP - flowPV;
                tmp_valveUnlim := accF + (2.0 + 0.5 * scanSeconds) * tmp_eF;
                valveCommand := LIMIT(0.0, tmp_valveUnlim, 100.0);

            2:
                tmp_eT := tempSP - tempPV;
                tmp_flowUnlim := accT + (1.0 + 0.2 * scanSeconds) * tmp_eT;
                flowSP := LIMIT(0.0, tmp_flowUnlim, 50.0);

                tmp_eF := flowSP - flowPV;
                tmp_valveUnlim := accF + (2.0 + 0.5 * scanSeconds) * tmp_eF;
                valveCommand := LIMIT(0.0, tmp_valveUnlim, 100.0);
        END_CASE;
    END_IF;
END_IF;

(* 用最终输出回算积分量，保证无扰切换和抗积分饱和 *)
tmp_eT := tempSP - tempPV;
tmp_eF := flowSP - flowPV;
accT := flowSP - 1.0 * tmp_eT;
accF := valveCommand - 2.0 * tmp_eF;

prevFlowSP := flowSP;
prevValveCmd := valveCommand;
prevMode := mode;
prevResetBtn := resetBtn;
first := FALSE;

END_FUNCTION_BLOCK

(* ---- self-hard-07.raw_candidate_01.st ---- *)
FUNCTION_BLOCK FB
VAR_INPUT
    mode : INT;
    resetBtn : BOOL;
    scanSeconds : REAL;
    tempSP : REAL;
    tempPV : REAL;
    flowPV : REAL;
    manualFlowSP : REAL;
    manualValve : REAL;
END_VAR
VAR_OUTPUT
    flowSP : REAL;
    valveCommand : REAL;
    fault : BOOL;
    normalMode : BOOL;
END_VAR
VAR
    first : BOOL := TRUE;
    prevMode : INT := 0;
    prevResetBtn : BOOL := FALSE;
    prevFlowSP : REAL := 0.0;
    prevValveCmd : REAL := 0.0;
    accT : REAL := 0.0;
    accF : REAL := 0.0;
    tmp_eT : REAL;
    tmp_eF : REAL;
    tmp_flowUnlim : REAL;
    tmp_valveUnlim : REAL;
    tmp_resetRising : BOOL;
    tmp_modeChanged : BOOL;
END_VAR

(* ENGINEERING_CONTRACT
   flowSP: manual/limited PI output; retained via prevFlowSP between scans; reset/fault/switch presets.
   valveCommand: manual/limited PI output; retained via prevValveCmd; reset/fault/switch presets.
   fault: combinational from mode/scanSeconds; no latch.
   normalMode: true only in stable valid mode with no first/reset/fault/mode change.
   Reset rising: outputs=manual values, integrators preloaded; fault still reports current mode/scanSeconds.
   PI back-calculates accT/accF from final outputs every scan, preventing integral windup.
   Units: flowSP t/h, valveCommand %, accT t/h, accF %, scanSeconds s. PUB001-PUB065.
*)
(* CONTRACT_RULES [] *)

fault := (mode < 0) OR (mode > 2) OR (scanSeconds <= 0.0) OR (scanSeconds > 10.0);
tmp_resetRising := resetBtn AND NOT prevResetBtn;
normalMode := FALSE;

IF first THEN
    flowSP := manualFlowSP;
    valveCommand := manualValve;
ELSIF fault THEN
    flowSP := manualFlowSP;
    valveCommand := manualValve;
ELSIF tmp_resetRising THEN
    flowSP := manualFlowSP;
    valveCommand := manualValve;
ELSE
    tmp_modeChanged := (mode <> prevMode);
    IF tmp_modeChanged THEN
        IF mode = 2 THEN
            flowSP := prevFlowSP;
            valveCommand := prevValveCmd;
        ELSE
            flowSP := manualFlowSP;
            valveCommand := prevValveCmd;
        END_IF;
    ELSE
        normalMode := TRUE;
        CASE mode OF
            0:
                flowSP := manualFlowSP;
                valveCommand := manualValve;

            1:
                flowSP := manualFlowSP;
                tmp_eF := flowSP - flowPV;
                tmp_valveUnlim := accF + (2.0 + 0.5 * scanSeconds) * tmp_eF;
                valveCommand := LIMIT(0.0, tmp_valveUnlim, 100.0);

            2:
                tmp_eT := tempSP - tempPV;
                tmp_flowUnlim := accT + (1.0 + 0.2 * scanSeconds) * tmp_eT;
                flowSP := LIMIT(0.0, tmp_flowUnlim, 50.0);

                tmp_eF := flowSP - flowPV;
                tmp_valveUnlim := accF + (2.0 + 0.5 * scanSeconds) * tmp_eF;
                valveCommand := LIMIT(0.0, tmp_valveUnlim, 100.0);
        END_CASE;
    END_IF;
END_IF;

(* 用最终输出回算积分量，保证无扰切换和抗积分饱和 *)
tmp_eT := tempSP - tempPV;
tmp_eF := flowSP - flowPV;
accT := flowSP - 1.0 * tmp_eT;
accF := valveCommand - 2.0 * tmp_eF;

prevFlowSP := flowSP;
prevValveCmd := valveCommand;
prevMode := mode;
prevResetBtn := resetBtn;
first := FALSE;

END_FUNCTION_BLOCK

(* ---- self-medium-01.candidate_01.st ---- *)
TYPE ST_Recipe :
STRUCT
    recipeID : INT;
    totalRatio : REAL;
    temperature : REAL;
END_STRUCT
END_TYPE;

(* ENGINEERING_CONTRACT
valid: set TRUE only on accepted load edge (loadCmd rising AND NOT running, slot 1..8, recipeID<>0, totalRatio 99..101, temperature 30..180). Set FALSE on accepted invalid edge. Otherwise retains latched value; initial FALSE.
loadedID: set to recipe[selSlot].recipeID on accepted valid edge. Set 0 on accepted invalid edge, including empty/out-of-range/ratio/temp. Retains latched value when no accepted edge or running=TRUE; initial 0.
Priority: running gates loading; no edge processing while running.
Edge: detected once per loadCmd false-to-true scan via local_prevLoadCmd.
Boundaries: inclusive REAL comparisons. Array access only after selSlot 1..8.
*)

(* CONTRACT_RULES [] *)

FUNCTION_BLOCK FB
VAR_INPUT
    recipe : ARRAY[1..8] OF ST_Recipe;
    selSlot : INT;
    loadCmd : BOOL;
    running : BOOL;
END_VAR
VAR_OUTPUT
    valid : BOOL;
    loadedID : INT;
END_VAR
VAR
    local_prevLoadCmd : BOOL := FALSE;
    local_edge : BOOL;
    local_slot : INT;
    local_latchedValid : BOOL := FALSE;
    local_latchedID : INT := 0;
END_VAR

local_edge := loadCmd AND NOT local_prevLoadCmd;
local_prevLoadCmd := loadCmd;

IF local_edge AND NOT running THEN
    local_slot := selSlot;
    IF (local_slot >= 1) AND (local_slot <= 8) THEN
        IF (recipe[local_slot].recipeID <> 0)
           AND (recipe[local_slot].totalRatio >= 99.0)
           AND (recipe[local_slot].totalRatio <= 101.0)
           AND (recipe[local_slot].temperature >= 30.0)
           AND (recipe[local_slot].temperature <= 180.0) THEN
            local_latchedValid := TRUE;
            local_latchedID := recipe[local_slot].recipeID;
        ELSE
            local_latchedValid := FALSE;
            local_latchedID := 0;
        END_IF;
    ELSE
        local_latchedValid := FALSE;
        local_latchedID := 0;
    END_IF;
END_IF;

valid := local_latchedValid;
loadedID := local_latchedID;

END_FUNCTION_BLOCK

(* ---- self-medium-01.raw_candidate_01.st ---- *)
TYPE ST_Recipe :
STRUCT
    recipeID : INT;
    totalRatio : REAL;
    temperature : REAL;
END_STRUCT
END_TYPE

(* ENGINEERING_CONTRACT
valid: set TRUE only on accepted load edge (loadCmd rising AND NOT running, slot 1..8, recipeID<>0, totalRatio 99..101, temperature 30..180). Set FALSE on accepted invalid edge. Otherwise retains latched value; initial FALSE.
loadedID: set to recipe[selSlot].recipeID on accepted valid edge. Set 0 on accepted invalid edge, including empty/out-of-range/ratio/temp. Retains latched value when no accepted edge or running=TRUE; initial 0.
Priority: running gates loading; no edge processing while running.
Edge: detected once per loadCmd false-to-true scan via local_prevLoadCmd.
Boundaries: inclusive REAL comparisons. Array access only after selSlot 1..8.
*)

(* CONTRACT_RULES [] *)

FUNCTION_BLOCK FB
VAR_INPUT
    recipe : ARRAY[1..8] OF ST_Recipe;
    selSlot : INT;
    loadCmd : BOOL;
    running : BOOL;
END_VAR
VAR_OUTPUT
    valid : BOOL;
    loadedID : INT;
END_VAR
VAR
    local_prevLoadCmd : BOOL := FALSE;
    local_edge : BOOL;
    local_slot : INT;
    local_latchedValid : BOOL := FALSE;
    local_latchedID : INT := 0;
END_VAR

local_edge := loadCmd AND NOT local_prevLoadCmd;
local_prevLoadCmd := loadCmd;

IF local_edge AND NOT running THEN
    local_slot := selSlot;
    IF (local_slot >= 1) AND (local_slot <= 8) THEN
        IF (recipe[local_slot].recipeID <> 0)
           AND (recipe[local_slot].totalRatio >= 99.0)
           AND (recipe[local_slot].totalRatio <= 101.0)
           AND (recipe[local_slot].temperature >= 30.0)
           AND (recipe[local_slot].temperature <= 180.0) THEN
            local_latchedValid := TRUE;
            local_latchedID := recipe[local_slot].recipeID;
        ELSE
            local_latchedValid := FALSE;
            local_latchedID := 0;
        END_IF;
    ELSE
        local_latchedValid := FALSE;
        local_latchedID := 0;
    END_IF;
END_IF;

valid := local_latchedValid;
loadedID := local_latchedID;

END_FUNCTION_BLOCK

(* ---- self-medium-02.candidate_01.st ---- *)
(*
ENGINEERING_CONTRACT
- filteredValue: combinational average of actual buffer samples while enable=TRUE; retained unchanged when enable=FALSE (PUB006/S5).
- windowFull: retained full flag; set TRUE when sampleCount reaches 8; held while enabled; reset only by enable=FALSE (PUB005/S2/S3).
- sampleCount: state; increments on each enabled scan up to 8; held at 8 while enabled; reset to 0 same scan on disable (PUB004/S3/S4).
- buffer: 8-slot ring; never zero-filled in average; partial count uses only actual samples PUB001/PUB002/S1; full count FIFO overwrite oldest PUB003.
- Priority: enable=FALSE clears history/window and leaves filteredValue untouched before any sampling.
- Units/boundaries: rawValue/filteredValue REAL sample units; sampleCount INT 0..8; threshold exactly 8.
*)
(* CONTRACT_RULES [] *)
FUNCTION_BLOCK FB
VAR_INPUT
    enable : BOOL;
    rawValue : REAL;
END_VAR
VAR_OUTPUT
    filteredValue : REAL;
    windowFull : BOOL;
    sampleCount : INT;
END_VAR
VAR
    tmp_buffer : ARRAY[0..7] OF REAL;
    tmp_count : INT := 0;
    tmp_head : INT := 0;
    tmp_i : INT;
    tmp_sum : REAL;
END_VAR

IF enable THEN
    tmp_buffer[tmp_head] := rawValue;
    tmp_head := ((tmp_head + 1) MOD 8);
    IF tmp_count < 8 THEN
        tmp_count := tmp_count + 1;
    END_IF;
    sampleCount := tmp_count;
    windowFull := (tmp_count >= 8);
    tmp_sum := 0.0;
    IF tmp_count > 0 THEN
        FOR tmp_i := 0 TO tmp_count - 1 DO
            tmp_sum := tmp_sum + tmp_buffer[tmp_i];
        END_FOR;
        filteredValue := tmp_sum / INT_TO_REAL(tmp_count);
    END_IF;
ELSE
    tmp_count := 0;
    tmp_head := 0;
    sampleCount := 0;
    windowFull := FALSE;
    FOR tmp_i := 0 TO 7 DO
        tmp_buffer[tmp_i] := 0.0;
    END_FOR;
    (* filteredValue intentionally remains at last computed result *)
END_IF;
END_FUNCTION_BLOCK

(* ---- self-medium-02.raw_candidate_01.st ---- *)
(*
ENGINEERING_CONTRACT
- filteredValue: combinational average of actual buffer samples while enable=TRUE; retained unchanged when enable=FALSE (PUB006/S5).
- windowFull: retained full flag; set TRUE when sampleCount reaches 8; held while enabled; reset only by enable=FALSE (PUB005/S2/S3).
- sampleCount: state; increments on each enabled scan up to 8; held at 8 while enabled; reset to 0 same scan on disable (PUB004/S3/S4).
- buffer: 8-slot ring; never zero-filled in average; partial count uses only actual samples PUB001/PUB002/S1; full count FIFO overwrite oldest PUB003.
- Priority: enable=FALSE clears history/window and leaves filteredValue untouched before any sampling.
- Units/boundaries: rawValue/filteredValue REAL sample units; sampleCount INT 0..8; threshold exactly 8.
*)
(* CONTRACT_RULES [] *)
FUNCTION_BLOCK FB
VAR_INPUT
    enable : BOOL;
    rawValue : REAL;
END_VAR
VAR_OUTPUT
    filteredValue : REAL;
    windowFull : BOOL;
    sampleCount : INT;
END_VAR
VAR
    tmp_buffer : ARRAY[0..7] OF REAL;
    tmp_count : INT := 0;
    tmp_head : INT := 0;
    tmp_i : INT;
    tmp_sum : REAL;
END_VAR

IF enable THEN
    tmp_buffer[tmp_head] := rawValue;
    tmp_head := ((tmp_head + 1) MOD 8);
    IF tmp_count < 8 THEN
        tmp_count := tmp_count + 1;
    END_IF;
    sampleCount := tmp_count;
    windowFull := (tmp_count >= 8);
    tmp_sum := 0.0;
    IF tmp_count > 0 THEN
        FOR tmp_i := 0 TO tmp_count - 1 DO
            tmp_sum := tmp_sum + tmp_buffer[tmp_i];
        END_FOR;
        filteredValue := tmp_sum / INT_TO_REAL(tmp_count);
    END_IF;
ELSE
    tmp_count := 0;
    tmp_head := 0;
    sampleCount := 0;
    windowFull := FALSE;
    FOR tmp_i := 0 TO 7 DO
        tmp_buffer[tmp_i] := 0.0;
    END_FOR;
    (* filteredValue intentionally remains at last computed result *)
END_IF;
END_FUNCTION_BLOCK

(* ---- self-medium-03.candidate_01.st ---- *)
FUNCTION_BLOCK FB
(* ENGINEERING_CONTRACT
   Output group motorUp/motorDown/errorFlag:
   - motorUp activation: state=OPENING while !obstacle and !openLimit (PUB003, PUB010, PUB012).
   - motorDown activation: state=CLOSING while !obstacle and !closeLimit (PUB003, PUB011, PUB013).
   - Retention: motion continues after button release until own limit, obstacle, or FAULT reset (PUB003, PUB012, PUB013).
   - Deactivation: own limit stops and returns to IDLE same scan; obstacle or FAULT stops both (PUB004-PUB006).
   - Same-scan priority: obstacle > limit/motion/reset; reset only returns to IDLE with motors stopped (PUB005, PUB007).
   - errorFlag activation: any obstacle, latched in FAULT (PUB004, PUB006).
   - errorFlag reset: only !obstacle and rising(openBtn AND closeBtn) (PUB007); no release-while-held auto reset.
   - Units/boundaries: BOOL signals; no timers; S1-S14 motor exclusion and latching contracts.
*)
(* CONTRACT_RULES [] *)
VAR_INPUT
    openBtn: BOOL;
    closeBtn: BOOL;
    openLimit: BOOL;
    closeLimit: BOOL;
    obstacle: BOOL;
END_VAR
VAR_OUTPUT
    motorUp: BOOL;
    motorDown: BOOL;
    errorFlag: BOOL;
END_VAR
VAR
    state: INT := 0; (* 0: IDLE, 1: OPENING, 2: CLOSING, 3: FAULT *)
    latchedFault: BOOL := FALSE;
    prevOpenBtn: BOOL := FALSE;
    prevCloseBtn: BOOL := FALSE;
    tmp_rOpen: BOOL;
    tmp_rClose: BOOL;
    tmp_rBoth: BOOL;
    tmp_state: INT;
    tmp_fault: BOOL;
    tmp_up: BOOL;
    tmp_down: BOOL;
END_VAR

tmp_rOpen := openBtn AND NOT prevOpenBtn;
tmp_rClose := closeBtn AND NOT prevCloseBtn;
tmp_rBoth := openBtn AND closeBtn AND NOT (prevOpenBtn AND prevCloseBtn);

tmp_state := state;
tmp_fault := latchedFault;
tmp_up := FALSE;
tmp_down := FALSE;

IF obstacle THEN
    tmp_state := 3;
    tmp_fault := TRUE;
ELSE
    IF state = 3 THEN
        IF tmp_rBoth THEN
            tmp_state := 0;
            tmp_fault := FALSE;
        END_IF;
    ELSIF state = 0 THEN
        IF tmp_rOpen AND NOT closeBtn AND NOT openLimit THEN
            tmp_state := 1;
            tmp_up := TRUE;
        ELSIF tmp_rClose AND NOT openBtn AND NOT closeLimit THEN
            tmp_state := 2;
            tmp_down := TRUE;
        END_IF;
    ELSIF state = 1 THEN
        IF openLimit THEN
            tmp_state := 0;
        ELSE
            tmp_up := TRUE;
        END_IF;
    ELSIF state = 2 THEN
        IF closeLimit THEN
            tmp_state := 0;
        ELSE
            tmp_down := TRUE;
        END_IF;
    END_IF;
END_IF;

state := tmp_state;
latchedFault := tmp_fault;
motorUp := tmp_up;
motorDown := tmp_down;
errorFlag := latchedFault;

prevOpenBtn := openBtn;
prevCloseBtn := closeBtn;

END_FUNCTION_BLOCK

(* ---- self-medium-03.raw_candidate_01.st ---- *)
FUNCTION_BLOCK FB
(* ENGINEERING_CONTRACT
   Output group motorUp/motorDown/errorFlag:
   - motorUp activation: state=OPENING while !obstacle and !openLimit (PUB003, PUB010, PUB012).
   - motorDown activation: state=CLOSING while !obstacle and !closeLimit (PUB003, PUB011, PUB013).
   - Retention: motion continues after button release until own limit, obstacle, or FAULT reset (PUB003, PUB012, PUB013).
   - Deactivation: own limit stops and returns to IDLE same scan; obstacle or FAULT stops both (PUB004-PUB006).
   - Same-scan priority: obstacle > limit/motion/reset; reset only returns to IDLE with motors stopped (PUB005, PUB007).
   - errorFlag activation: any obstacle, latched in FAULT (PUB004, PUB006).
   - errorFlag reset: only !obstacle and rising(openBtn AND closeBtn) (PUB007); no release-while-held auto reset.
   - Units/boundaries: BOOL signals; no timers; S1-S14 motor exclusion and latching contracts.
*)
(* CONTRACT_RULES [] *)
VAR_INPUT
    openBtn: BOOL;
    closeBtn: BOOL;
    openLimit: BOOL;
    closeLimit: BOOL;
    obstacle: BOOL;
END_VAR
VAR_OUTPUT
    motorUp: BOOL;
    motorDown: BOOL;
    errorFlag: BOOL;
END_VAR
VAR
    state: INT := 0; (* 0: IDLE, 1: OPENING, 2: CLOSING, 3: FAULT *)
    latchedFault: BOOL := FALSE;
    prevOpenBtn: BOOL := FALSE;
    prevCloseBtn: BOOL := FALSE;
    tmp_rOpen: BOOL;
    tmp_rClose: BOOL;
    tmp_rBoth: BOOL;
    tmp_state: INT;
    tmp_fault: BOOL;
    tmp_up: BOOL;
    tmp_down: BOOL;
END_VAR

tmp_rOpen := openBtn AND NOT prevOpenBtn;
tmp_rClose := closeBtn AND NOT prevCloseBtn;
tmp_rBoth := openBtn AND closeBtn AND NOT (prevOpenBtn AND prevCloseBtn);

tmp_state := state;
tmp_fault := latchedFault;
tmp_up := FALSE;
tmp_down := FALSE;

IF obstacle THEN
    tmp_state := 3;
    tmp_fault := TRUE;
ELSE
    IF state = 3 THEN
        IF tmp_rBoth THEN
            tmp_state := 0;
            tmp_fault := FALSE;
        END_IF
    ELSIF state = 0 THEN
        IF tmp_rOpen AND NOT closeBtn AND NOT openLimit THEN
            tmp_state := 1;
            tmp_up := TRUE;
        ELSIF tmp_rClose AND NOT openBtn AND NOT closeLimit THEN
            tmp_state := 2;
            tmp_down := TRUE;
        END_IF
    ELSIF state = 1 THEN
        IF openLimit THEN
            tmp_state := 0;
        ELSE
            tmp_up := TRUE;
        END_IF
    ELSIF state = 2 THEN
        IF closeLimit THEN
            tmp_state := 0;
        ELSE
            tmp_down := TRUE;
        END_IF
    END_IF
END_IF

state := tmp_state;
latchedFault := tmp_fault;
motorUp := tmp_up;
motorDown := tmp_down;
errorFlag := latchedFault;

prevOpenBtn := openBtn;
prevCloseBtn := closeBtn;

END_FUNCTION_BLOCK

(* ---- self-medium-04.candidate_01.st ---- *)
(* ENGINEERING_CONTRACT
- valveOpen: set TRUE only by start edge from idle/pending; held while filling below target; set FALSE same scan when accum>=target or reset edge. Same-scan reset priority over start/flow/confirm. S2,S7,S8,S9,S12,S13.
- fillsToday: increments once only when local_pending AND doneSensor; reset edge zeroes same scan; saturates at 32767 while still clearing local_pending. S1,S3,S4,S6,S10,S11,S14.
- local_pending: set when threshold reached; cleared by confirm, reset, or start-new-bottle cancellation. S4,S10,S11,S13,S14.
- local_accum: cleared by reset/start; adds flowVol only while local_filling including start scan; compare >= targetVol. S5,S8,S12.
- local_filling: filling process state; start edge activates; threshold/reset deactivates.
- Edge memory false before first call; doneSensor read as level. Units: volume REAL mL, count INT max 32767.
*)
(* CONTRACT_RULES [] *)
FUNCTION_BLOCK FB
VAR_INPUT
    startBtn : BOOL;
    resetBtn : BOOL;
    doneSensor : BOOL;
    targetVol : REAL;
    flowVol : REAL;
END_VAR
VAR_OUTPUT
    valveOpen : BOOL := FALSE;
    fillsToday : INT := 0;
END_VAR
VAR
    tmp_prevStart : BOOL := FALSE;
    tmp_prevReset : BOOL := FALSE;
    local_accum : REAL := 0.0;
    local_filling : BOOL := FALSE;
    local_pending : BOOL := FALSE;
    local_startR : BOOL;
    local_resetR : BOOL;
END_VAR

local_startR := startBtn AND (NOT tmp_prevStart);
local_resetR := resetBtn AND (NOT tmp_prevReset);

IF local_resetR THEN
    valveOpen := FALSE;
    fillsToday := 0;
    local_accum := 0.0;
    local_filling := FALSE;
    local_pending := FALSE;
ELSE
    IF local_startR AND (NOT local_filling) THEN
        local_pending := FALSE;
        local_filling := TRUE;
        valveOpen := TRUE;
        local_accum := 0.0;
    END_IF;

    IF local_filling THEN
        local_accum := local_accum + flowVol;
        IF local_accum >= targetVol THEN
            local_filling := FALSE;
            valveOpen := FALSE;
            local_pending := TRUE;
        END_IF;
    END_IF;

    IF local_pending AND doneSensor THEN
        IF fillsToday < 32767 THEN
            fillsToday := fillsToday + 1;
        END_IF;
        local_pending := FALSE;
    END_IF;
END_IF;

tmp_prevStart := startBtn;
tmp_prevReset := resetBtn;
END_FUNCTION_BLOCK

(* ---- self-medium-04.raw_candidate_01.st ---- *)
(* ENGINEERING_CONTRACT
- valveOpen: set TRUE only by start edge from idle/pending; held while filling below target; set FALSE same scan when accum>=target or reset edge. Same-scan reset priority over start/flow/confirm. S2,S7,S8,S9,S12,S13.
- fillsToday: increments once only when local_pending AND doneSensor; reset edge zeroes same scan; saturates at 32767 while still clearing local_pending. S1,S3,S4,S6,S10,S11,S14.
- local_pending: set when threshold reached; cleared by confirm, reset, or start-new-bottle cancellation. S4,S10,S11,S13,S14.
- local_accum: cleared by reset/start; adds flowVol only while local_filling including start scan; compare >= targetVol. S5,S8,S12.
- local_filling: filling process state; start edge activates; threshold/reset deactivates.
- Edge memory false before first call; doneSensor read as level. Units: volume REAL mL, count INT max 32767.
*)
(* CONTRACT_RULES [] *)
FUNCTION_BLOCK FB
VAR_INPUT
    startBtn : BOOL;
    resetBtn : BOOL;
    doneSensor : BOOL;
    targetVol : REAL;
    flowVol : REAL;
END_VAR
VAR_OUTPUT
    valveOpen : BOOL := FALSE;
    fillsToday : INT := 0;
END_VAR
VAR
    tmp_prevStart : BOOL := FALSE;
    tmp_prevReset : BOOL := FALSE;
    local_accum : REAL := 0.0;
    local_filling : BOOL := FALSE;
    local_pending : BOOL := FALSE;
    local_startR : BOOL;
    local_resetR : BOOL;
END_VAR

local_startR := startBtn AND (NOT tmp_prevStart);
local_resetR := resetBtn AND (NOT tmp_prevReset);

IF local_resetR THEN
    valveOpen := FALSE;
    fillsToday := 0;
    local_accum := 0.0;
    local_filling := FALSE;
    local_pending := FALSE;
ELSE
    IF local_startR AND (NOT local_filling) THEN
        local_pending := FALSE;
        local_filling := TRUE;
        valveOpen := TRUE;
        local_accum := 0.0;
    END_IF;

    IF local_filling THEN
        local_accum := local_accum + flowVol;
        IF local_accum >= targetVol THEN
            local_filling := FALSE;
            valveOpen := FALSE;
            local_pending := TRUE;
        END_IF;
    END_IF;

    IF local_pending AND doneSensor THEN
        IF fillsToday < 32767 THEN
            fillsToday := fillsToday + 1;
        END_IF;
        local_pending := FALSE;
    END_IF;
END_IF;

tmp_prevStart := startBtn;
tmp_prevReset := resetBtn;
END_FUNCTION_BLOCK

(* ---- self-medium-05.candidate_01.st ---- *)
FUNCTION_BLOCK FB
VAR_INPUT
    enable : BOOL;
    resetBtn : BOOL;
    scanSeconds : LREAL;
    steamFlow : LREAL;
    fuelFlow : LREAL;
    steamTemp : LREAL;
    steamPressure : LREAL;
END_VAR
VAR_OUTPUT
    qualified : BOOL;
    dataFault : BOOL;
    qualifiedTon : LREAL;
    fuelTon : LREAL;
    revenue : LREAL;
    cost : LREAL;
    netProfit : LREAL;
END_VAR
VAR
    lastResetBtn : BOOL := FALSE;
    tmp_resetRising : BOOL;
END_VAR

(* ENGINEERING_CONTRACT
   qualified: combinational per PUB001-S1, ranges closed.
   dataFault: combinational per PUB004, bounds scanSeconds/(0,10], steamFlow [0,90], fuelFlow [0,6].
   qualifiedTon: retained accum; reset on rising resetBtn to 0 same scan; priority over fault/disable.
   fuelTon: retained accum; reset same rising edge; priority over fault/disable.
   revenue/cost/netProfit: derived each scan from tonnage*unit price; money units CNY.
   Reset rising: resetBtn AND NOT lastResetBtn; first TRUE scan counted; held TRUE no repeat.
   Non-negative accum guaranteed by valid inputs and reset; netProfit may be negative.
*)

(* CONTRACT_RULES [] *)

tmp_resetRising := resetBtn AND NOT lastResetBtn;

qualified := (steamTemp >= 447.0) AND (steamTemp <= 453.0)
             AND (steamPressure >= 3750.0) AND (steamPressure <= 3850.0);

dataFault := (scanSeconds <= 0.0) OR (scanSeconds > 10.0)
             OR (steamFlow < 0.0) OR (steamFlow > 90.0)
             OR (fuelFlow < 0.0) OR (fuelFlow > 6.0);

IF tmp_resetRising THEN
    qualifiedTon := 0.0;
    fuelTon := 0.0;
ELSE
    IF enable AND NOT dataFault THEN
        fuelTon := fuelTon + (fuelFlow * scanSeconds / 1000.0);
        IF qualified THEN
            qualifiedTon := qualifiedTon + (steamFlow * scanSeconds / 1000.0);
        END_IF;
    END_IF;
END_IF;

revenue := qualifiedTon * 280.0;
cost := fuelTon * 1500.0;
netProfit := revenue - cost;

lastResetBtn := resetBtn;

END_FUNCTION_BLOCK

(* ---- self-medium-05.raw_candidate_01.st ---- *)
FUNCTION_BLOCK FB
VAR_INPUT
    enable : BOOL;
    resetBtn : BOOL;
    scanSeconds : LREAL;
    steamFlow : LREAL;
    fuelFlow : LREAL;
    steamTemp : LREAL;
    steamPressure : LREAL;
END_VAR
VAR_OUTPUT
    qualified : BOOL;
    dataFault : BOOL;
    qualifiedTon : LREAL;
    fuelTon : LREAL;
    revenue : LREAL;
    cost : LREAL;
    netProfit : LREAL;
END_VAR
VAR
    lastResetBtn : BOOL := FALSE;
    tmp_resetRising : BOOL;
END_VAR

(* ENGINEERING_CONTRACT
   qualified: combinational per PUB001-S1, ranges closed.
   dataFault: combinational per PUB004, bounds scanSeconds/(0,10], steamFlow [0,90], fuelFlow [0,6].
   qualifiedTon: retained accum; reset on rising resetBtn to 0 same scan; priority over fault/disable.
   fuelTon: retained accum; reset same rising edge; priority over fault/disable.
   revenue/cost/netProfit: derived each scan from tonnage*unit price; money units CNY.
   Reset rising: resetBtn AND NOT lastResetBtn; first TRUE scan counted; held TRUE no repeat.
   Non-negative accum guaranteed by valid inputs and reset; netProfit may be negative.
*)

(* CONTRACT_RULES [] *)

tmp_resetRising := resetBtn AND NOT lastResetBtn;

qualified := (steamTemp >= 447.0) AND (steamTemp <= 453.0)
             AND (steamPressure >= 3750.0) AND (steamPressure <= 3850.0);

dataFault := (scanSeconds <= 0.0) OR (scanSeconds > 10.0)
             OR (steamFlow < 0.0) OR (steamFlow > 90.0)
             OR (fuelFlow < 0.0) OR (fuelFlow > 6.0);

IF tmp_resetRising THEN
    qualifiedTon := 0.0;
    fuelTon := 0.0;
ELSE
    IF enable AND NOT dataFault THEN
        fuelTon := fuelTon + (fuelFlow * scanSeconds / 1000.0);
        IF qualified THEN
            qualifiedTon := qualifiedTon + (steamFlow * scanSeconds / 1000.0);
        END_IF;
    END_IF;
END_IF;

revenue := qualifiedTon * 280.0;
cost := fuelTon * 1500.0;
netProfit := revenue - cost;

lastResetBtn := resetBtn;

END_FUNCTION_BLOCK

(* ---- self-medium-06.candidate_01.st ---- *)
FUNCTION_BLOCK FB
VAR_INPUT
    enable: BOOL;
    resetBtn: BOOL;
    sensorValid: BOOL;
    setpoint: REAL;
    temperature: REAL;
    scanSeconds: REAL;
    bias: REAL;
END_VAR
VAR_OUTPUT
    power: REAL;
    correction: REAL;
    fault: BOOL;
END_VAR
VAR
    ePrev: REAL := 0.0;
    histValid: BOOL := FALSE;
    resetRTrig: R_TRIG;
    resetEdge: BOOL;
    e: REAL;
    x: REAL;
    y: REAL;
    de: REAL;
END_VAR

(* ENGINEERING_CONTRACT
   - fault (PUB004/PUB032/S4): combinational from sensorValid and scanSeconds; no retention; updated every scan.
   - power/correction: combinational outputs from current inputs and internal history; not latched except zero-clear on !enable/fault/reset rise.
   - Clear on !enable OR fault OR resetBtn rising edge (PUB005): same scan, zero outputs and clear history (ePrev=0, histValid=false); reset edge is one-shot.
   - Valid first/cleared-history scan (PUB005): de=0, correction=20*clamp(e/10, -1, 1); equivalent to y=0.
   - Valid with previous history (PUB004/PUB006): de=(e-ePrev)/scanSeconds; y=clamp(de/2,-1,1); correction=20*x+10*y (S13 equivalence).
   - power = LIMIT(0, bias+correction, 100) (PUB005/S1/S10); correction within ±30 by construction.
   - Units: temp °C, scan seconds s, bias/power/correction %, e/10 and de/2 dimensionless.
   - History update: after any valid computation, ePrev=e, histValid=true; otherwise reset.
   - Same-scan priority: clear condition dominates computation.
*)
(* CONTRACT_RULES [] *)

fault := (NOT sensorValid) OR (scanSeconds <= 0.0) OR (scanSeconds > 10.0);

resetRTrig(CLK := resetBtn);
resetEdge := resetRTrig.Q;

IF (NOT enable) OR fault OR resetEdge THEN
    power := 0.0;
    correction := 0.0;
    ePrev := 0.0;
    histValid := FALSE;
ELSE
    e := setpoint - temperature;
    x := LIMIT(-1.0, e / 10.0, 1.0);

    IF NOT histValid THEN
        de := 0.0;
        y := 0.0;
        correction := 20.0 * x;
    ELSE
        de := (e - ePrev) / scanSeconds;
        y := LIMIT(-1.0, de / 2.0, 1.0);
        correction := 20.0 * x + 10.0 * y;
    END_IF;

    power := LIMIT(0.0, bias + correction, 100.0);

    histValid := TRUE;
    ePrev := e;
END_IF;

END_FUNCTION_BLOCK

(* ---- self-medium-06.raw_candidate_01.st ---- *)
FUNCTION_BLOCK FB
VAR_INPUT
    enable: BOOL;
    resetBtn: BOOL;
    sensorValid: BOOL;
    setpoint: REAL;
    temperature: REAL;
    scanSeconds: REAL;
    bias: REAL;
END_VAR
VAR_OUTPUT
    power: REAL;
    correction: REAL;
    fault: BOOL;
END_VAR
VAR
    ePrev: REAL := 0.0;
    histValid: BOOL := FALSE;
    resetRTrig: R_TRIG;
    resetEdge: BOOL;
    e: REAL;
    x: REAL;
    y: REAL;
    de: REAL;
END_VAR

(* ENGINEERING_CONTRACT
   - fault (PUB004/PUB032/S4): combinational from sensorValid and scanSeconds; no retention; updated every scan.
   - power/correction: combinational outputs from current inputs and internal history; not latched except zero-clear on !enable/fault/reset rise.
   - Clear on !enable OR fault OR resetBtn rising edge (PUB005): same scan, zero outputs and clear history (ePrev=0, histValid=false); reset edge is one-shot.
   - Valid first/cleared-history scan (PUB005): de=0, correction=20*clamp(e/10, -1, 1); equivalent to y=0.
   - Valid with previous history (PUB004/PUB006): de=(e-ePrev)/scanSeconds; y=clamp(de/2,-1,1); correction=20*x+10*y (S13 equivalence).
   - power = LIMIT(0, bias+correction, 100) (PUB005/S1/S10); correction within ±30 by construction.
   - Units: temp °C, scan seconds s, bias/power/correction %, e/10 and de/2 dimensionless.
   - History update: after any valid computation, ePrev=e, histValid=true; otherwise reset.
   - Same-scan priority: clear condition dominates computation.
*)
(* CONTRACT_RULES [] *)

fault := (NOT sensorValid) OR (scanSeconds <= 0.0) OR (scanSeconds > 10.0);

resetRTrig(CLK := resetBtn);
resetEdge := resetRTrig.Q;

IF (NOT enable) OR fault OR resetEdge THEN
    power := 0.0;
    correction := 0.0;
    ePrev := 0.0;
    histValid := FALSE;
ELSE
    e := setpoint - temperature;
    x := LIMIT(-1.0, e / 10.0, 1.0);

    IF NOT histValid THEN
        de := 0.0;
        y := 0.0;
        correction := 20.0 * x;
    ELSE
        de := (e - ePrev) / scanSeconds;
        y := LIMIT(-1.0, de / 2.0, 1.0);
        correction := 20.0 * x + 10.0 * y;
    END_IF;

    power := LIMIT(0.0, bias + correction, 100.0);

    histValid := TRUE;
    ePrev := e;
END_IF;

END_FUNCTION_BLOCK
